// TIA Portal V20 export
// export: Created 2026-10-20T18:55:42.8916793Z, ExportSetting None, DisplayName Totally Integrated Automation Portal, DisplayVersion V20 Update 6, DisplayName TIA Portal Openness, DisplayVersion V20 Update 6, DisplayName TIA Portal Version Control Interface, DisplayVersion V20 Update 6, DisplayName SINAMICS Startdrive Advanced, DisplayVersion V20 SP1, DisplayName SINAMICS Startdrive G130, G150, S120, S150, SINAMICS MV, G220, S200, S210, DisplayVersion V20 SP1, DisplayName SINAMICS Startdrive G110M, G120, G120C, G120D, G120P, G115D, DisplayVersion V20 SP1, DisplayName STEP 7 Professional, DisplayVersion V20 Update 6, DisplayName STEP 7 Safety, DisplayVersion V20 Update 2, DisplayName WinCC Basic/Comfort/Advanced, DisplayVersion V20 Update 6, DisplayName WinCC Unified, DisplayVersion V20 Update 6
VAR_GLOBAL   // PLC tag table "Lock_2"
   Lamps_2 AT %QB880 : Byte;
   Lock_2_Estop_CH1 AT %I1766.2 : Bool;
   Lock_2_Closed_CH2 AT %I1766.1 : Bool;
   Switches_2 AT %IB299 : Byte;
   "Solenoid Enable_2" AT %Q881.0 : Bool;
   Lock_2_Estop_CH2 AT %I1766.3 : Bool;
   "Lock Reset_2" AT %Q1065.0 : Bool;
   Lock_2_Closed_CH1 AT %I1766.0 : Bool;
   Lock_2_Reset_Input2 AT %Q1767.1 : Bool;
   Lock_2_Reset_Input1 AT %Q1767.0 : Bool;
   Lock_2_Reset_Input3 AT %Q1767.2 : Bool;
   Lock_2_Reset_Input4 AT %Q1767.3 : Bool;
   "Lock Position_2" AT %I901.0 : Bool;
   "Guard Position_2" AT %I900.0 : Bool;
END_VAR
